(* PLC project Boiler_Control, CODESYS CODESYS V3.5 SP19 *)
(* stored: creationDateTime 2026-09-01T08:00:00 *)

PROGRAM PLC_PRG
  VAR
    TempSet : REAL;
  END_VAR

TempSet := 80.0;
END_PROGRAM

FUNCTION_BLOCK FB_Burner

END_FUNCTION_BLOCK

FUNCTION F_Scale


END_FUNCTION

CONFIGURATION Boiler_PLC
  RESOURCE Application ON PLC
    TASK MainTask(INTERVAL := T#20ms, PRIORITY := 1);
  END_RESOURCE
END_CONFIGURATION
